(* IEC 61131-3 sources: TcAgent_Knowledge/skills/plc-st-patterns/references, 8 files *)

(* ---- async_call.st ---- *)
/// Drives an asynchronous job with Execute, Busy, Done and Error: one edge per job, the result is kept until the next start.
/// Connect Execute to the block that does the job, and feed its Busy and Error back.
FUNCTION_BLOCK FB_AsyncCall
VAR_INPUT
	/// Starts a job on a rising edge
	Start : BOOL;
	/// Busy output of the called block
	JobBusy : BOOL;
	/// Error output of the called block
	JobError : BOOL;
	/// Longest time for a job
	Timeout : TIME;
END_VAR
VAR_OUTPUT
	/// To the Execute input of the called block
	Execute : BOOL;
	/// Job finished without an error
	Done : BOOL;
	/// Job failed or took too long
	Error : BOOL;
END_VAR
VAR
	_edge : R_TRIG;
	_timer : TON;
	_state : INT;
END_VAR
VAR CONSTANT
	STATE_IDLE : INT := 0;
	STATE_START : INT := 10;
	STATE_WAIT : INT := 20;
END_VAR
// --- implementation ---
_edge(CLK := Start);
_timer(IN := _state <> STATE_IDLE, PT := Timeout);

CASE _state OF
	STATE_IDLE:
		Execute := FALSE;
		IF _edge.Q THEN
			Done := FALSE;
			Error := FALSE;
			Execute := TRUE;
			_state := STATE_START;
		END_IF

	STATE_START:
		// the block needs one call with Execute before Busy can rise
		IF JobBusy THEN
			_state := STATE_WAIT;
		ELSIF JobError THEN
			Error := TRUE;
			_state := STATE_IDLE;
		ELSIF _timer.Q THEN
			Error := TRUE;
			_state := STATE_IDLE;
		END_IF

	STATE_WAIT:
		IF NOT JobBusy THEN
			Done := NOT JobError;
			Error := JobError;
			_state := STATE_IDLE;
		ELSIF _timer.Q THEN
			Error := TRUE;
			_state := STATE_IDLE;
		END_IF

ELSE
	Error := TRUE;
	_state := STATE_IDLE;
END_CASE

(* ---- debounce.st ---- *)
/// Debounces an input: the output follows only after the input was stable for the set time.
FUNCTION_BLOCK FB_Debounce
VAR_INPUT
	/// Raw input
	Raw : BOOL;
	/// How long the input must be stable
	Delay : TIME;
END_VAR
VAR_OUTPUT
	/// Debounced value
	Stable : BOOL;
END_VAR
VAR
	_on : TON;
	_off : TON;
END_VAR
// --- implementation ---
_on(IN := Raw, PT := Delay);
_off(IN := NOT Raw, PT := Delay);
IF _on.Q THEN
	Stable := TRUE;
ELSIF _off.Q THEN
	Stable := FALSE;
END_IF

(* ---- edge_counter.st ---- *)
/// Counts rising edges up to MaxCount; Reset has priority.
FUNCTION_BLOCK FB_EdgeCounter
VAR_INPUT
	/// Counted signal
	Pulse : BOOL;
	/// Sets the count to 0
	Reset : BOOL;
	/// Count at which Reached becomes TRUE (not "Limit": LIMIT is a standard function)
	MaxCount : UDINT;
END_VAR
VAR_OUTPUT
	/// Current count
	Count : UDINT;
	/// Count has reached MaxCount
	Reached : BOOL;
END_VAR
VAR
	_edge : R_TRIG;
END_VAR
// --- implementation ---
_edge(CLK := Pulse);
IF Reset THEN
	Count := 0;
ELSIF _edge.Q AND (Count < MaxCount) THEN
	Count := Count + 1;
END_IF
Reached := Count >= MaxCount;

(* ---- hysteresis.st ---- *)
/// Two-point control: on below Low, off above High, between them the state stays.
FUNCTION_BLOCK FB_Hysteresis
VAR_INPUT
	/// Measured value
	Value : LREAL;
	/// Switch on below this value
	Low : LREAL;
	/// Switch off above this value
	High : LREAL;
	/// FALSE switches off at once
	Enable : BOOL;
END_VAR
VAR_OUTPUT
	/// The output is on
	Active : BOOL;
	/// Low is not below High: the output stays off
	ConfigError : BOOL;
END_VAR
// --- implementation ---
ConfigError := Low >= High;
IF NOT Enable OR ConfigError THEN
	Active := FALSE;
ELSIF Value < Low THEN
	Active := TRUE;
ELSIF Value > High THEN
	Active := FALSE;
END_IF

(* ---- latch_priority.st ---- *)
/// Start/stop latch: stop has priority over start.
FUNCTION_BLOCK FB_LatchPriority
VAR_INPUT
	/// Start request
	Start : BOOL;
	/// TRUE = running allowed; FALSE stops, also on a broken wire
	StopOk : BOOL;
END_VAR
VAR_OUTPUT
	/// The output is on
	Running : BOOL;
END_VAR
// --- implementation ---
Running := StopOk AND (Start OR Running);

(* ---- shift_register.st ---- *)
/// Tracks parts on a conveyor: one position per clock edge, the state of each part travels with it.
FUNCTION_BLOCK FB_ShiftRegister
VAR_INPUT
	/// One edge per position of the conveyor
	Clock : BOOL;
	/// State of the part entering at position 1: 0 = none, 1 = good, 2 = bad
	InState : USINT;
	/// Clears all positions
	Clear : BOOL;
END_VAR
VAR_OUTPUT
	/// State of the part at each position
	Positions : ARRAY[1..LENGTH] OF USINT;
	/// State of the part that left at the last edge
	OutState : USINT;
END_VAR
VAR
	_edge : R_TRIG;
	_index : INT;
END_VAR
VAR CONSTANT
	LENGTH : INT := 8;
END_VAR
// --- implementation ---
_edge(CLK := Clock);
IF Clear THEN
	FOR _index := 1 TO LENGTH DO
		Positions[_index] := 0;
	END_FOR
	OutState := 0;
ELSIF _edge.Q THEN
	OutState := Positions[LENGTH];
	FOR _index := LENGTH TO 2 BY -1 DO
		Positions[_index] := Positions[_index - 1];
	END_FOR
	Positions[1] := InState;
END_IF

(* ---- timed_sequence.st ---- *)
/// Step sequence with a timeout per step and an error state that every step can reach.
FUNCTION_BLOCK FB_TimedSequence
VAR_INPUT
	/// Starts the sequence from Idle
	Start : BOOL;
	/// Acknowledges an error
	Reset : BOOL;
	/// Feedback: position reached
	AtWork : BOOL;
	/// Feedback: back in the start position
	AtHome : BOOL;
	/// Longest time per step
	StepTimeout : TIME;
END_VAR
VAR_OUTPUT
	/// Drive to the work position
	MoveToWork : BOOL;
	/// Drive back
	MoveToHome : BOOL;
	/// Sequence has stopped with an error
	Error : BOOL;
	/// Current step, for diagnosis
	Step : INT;
END_VAR
VAR
	_timer : TON;
	_lastStep : INT;
END_VAR
VAR CONSTANT
	STEP_IDLE : INT := 0;
	STEP_TO_WORK : INT := 10;
	STEP_TO_HOME : INT := 20;
	STEP_ERROR : INT := 900;
END_VAR
// --- implementation ---
// the timer runs anew in every step
_timer(IN := (Step = _lastStep) AND (Step <> STEP_IDLE) AND (Step <> STEP_ERROR), PT := StepTimeout);
_lastStep := Step;
MoveToWork := FALSE;
MoveToHome := FALSE;

CASE Step OF
	STEP_IDLE:
		IF Start THEN
			Step := STEP_TO_WORK;
		END_IF

	STEP_TO_WORK:
		MoveToWork := TRUE;
		IF AtWork THEN
			Step := STEP_TO_HOME;
		ELSIF _timer.Q THEN
			Step := STEP_ERROR;
		END_IF

	STEP_TO_HOME:
		MoveToHome := TRUE;
		IF AtHome THEN
			Step := STEP_IDLE;
		ELSIF _timer.Q THEN
			Step := STEP_ERROR;
		END_IF

	STEP_ERROR:
		IF Reset THEN
			Step := STEP_IDLE;
		END_IF

ELSE
	Step := STEP_ERROR;
END_CASE

Error := Step = STEP_ERROR;

(* ---- wait_timeout.st ---- *)
/// Waits for a signal with a timeout. Call it every cycle while Enable is TRUE.
FUNCTION_BLOCK FB_WaitTimeout
VAR_INPUT
	/// TRUE while waiting; FALSE resets
	Enable : BOOL;
	/// The awaited signal
	Signal : BOOL;
	/// Longest waiting time
	Timeout : TIME;
END_VAR
VAR_OUTPUT
	/// The signal came in time
	Done : BOOL;
	/// The signal did not come in time
	TimedOut : BOOL;
END_VAR
VAR
	_timer : TON;
END_VAR
// --- implementation ---
_timer(IN := Enable AND NOT Done, PT := Timeout);
IF NOT Enable THEN
	Done := FALSE;
	TimedOut := FALSE;
ELSIF NOT TimedOut THEN
	IF Signal THEN
		Done := TRUE;
	ELSIF _timer.Q THEN
		TimedOut := TRUE;
	END_IF
END_IF
